Staubli VAL3: utButton.pjx

--- utButton.pjx ---
Parameters version=s8.8.3Cs9_BS1660 stackSize=5000 millimeterUnit=true
Program file=start.pgx
Program file=stop.pgx
Data file=utButton.dtx
Type name=utAppearance path=./utAppearance/utAppearance.pjx
Type name=utBorder path=./utBorder/utBorder.pjx
Type name=utCommon path=./utCommon/utCommon.pjx
Type name=utText path=./utText/utText.pjx
Type name=utEvents path=./utEvents/utEvents.pjx
Type name=utData path=./utData/utData.pjx

--- utButton.dtx ---
public utAppearance Appearance
  [0]
    string sBackgroundColour
    string sBackgroundImage
    string sColour
    bool bVisibility
public utBorder Border
  [0]
    string sBorderColour
public utCommon Common
  [0]
    bool bDisabled
    string sText
    string sID
    string sPage
public utText Text
  [0]
    string sFontFamily
    string sFontStyle
    string sFontWeight
    string sTextAlignment
    num nFontSize
public utEvents Events
  [0]
    bool bClick
    bool bMouseDown
    bool bMouseUp
public utData Data
  [0]
    num nVal
    bool bStatus

--- start.pgx ---
program start()
begin
end

--- stop.pgx ---
program stop()
begin
end
